// TIA Portal V20 export
Screen "Robot_PLP_Kuka"  1276x673
  ScreenItem "Zone01" at 710,47 size 522x643  Type=HmiGraphicView
  ScreenItem "Rectangle TG Control" at 241,104 size 465x354  Type=HmiRectangle
  ScreenItem "permanentareaborderrectangle" at 0,0 size 0x0  Type=HmiRectangle
  ScreenItem "Line_Header_X0_Y64" at 0,64 size 1280x0  Type=HmiLine
  ScreenItem "nbgMessages" at 19,459 size 687x203  Type=HmiAlarmControl
  ScreenItem "Button_Back" at 2,2 size 90x60  Type=HmiButton
  ScreenItem "Rectangle Robot Status" at 19,104 size 222x354  Type=HmiRectangle
  ScreenItem "Text Filed E- Stop" at 129,207 size 100x21  Type=HmiTextBox
  ScreenItem "Text Field In Auto On" at 24,138 size 100x21  Type=HmiTextBox
  ScreenItem "Text Field Home Position" at 24,161 size 100x21  Type=HmiTextBox
  ScreenItem "Text field PLP Status" at 19,103 size 222x31  Type=HmiTextBox
  ScreenItem "Text Field Manual" at 129,138 size 100x21  Type=HmiTextBox
  ScreenItem "Text Field System Ready" at 24,184 size 100x21  Type=HmiTextBox
  ScreenItem "Text Field Motor On" at 24,207 size 100x21  Type=HmiTextBox
  ScreenItem "Text Field In Cycle" at 24,230 size 100x21  Type=HmiTextBox
  ScreenItem "Text Field Cycle On" at 24,253 size 100x21  Type=HmiTextBox
  ScreenItem "Text Field On Path" at 24,276 size 100x21  Type=HmiTextBox
  ScreenItem "Text Field ProgNumReq" at 24,299 size 100x21  Type=HmiTextBox
  ScreenItem "Text Field Task OK" at 24,322 size 100x21  Type=HmiTextBox
  ScreenItem "Text Field Tryout Mode" at 129,161 size 100x21  Type=HmiTextBox
  ScreenItem "Text Field Stop" at 129,184 size 100x21  Type=HmiTextBox
  ScreenItem "Text Filed Error" at 129,230 size 100x21  Type=HmiTextBox
  ScreenItem "IO Field Feedback Program" at 129,280 size 100x21  Type=HmiIOField
  ScreenItem "Text Field Feedback Program" at 134,250 size 89x30  Type=HmiTextBox
  ScreenItem "Text Field In Home Pos" at 24,345 size 100x21  Type=HmiTextBox
  ScreenItem "Text Field In Work Pos" at 24,368 size 100x21  Type=HmiTextBox
  ScreenItem "Text Field In Pounce Pos" at 24,391 size 100x21  Type=HmiTextBox
  ScreenItem "Rectangle Clear Style" at 251,262 size 85x56  Type=HmiRectangle
  ScreenItem "Button Clear Style" at 252,263 size 83x54  Type=HmiButton
  ScreenItem "Clear Style Interlock" at 0,0 size 100x30  Type=HmiCircle
  ScreenItem "Rectangle Select Style1" at 251,140 size 85x56  Type=HmiRectangle
  ScreenItem "Button Select Style1" at 252,141 size 83x54  Type=HmiButton
  ScreenItem "Select Style Interlock1" at 0,0 size 100x30  Type=HmiCircle
  ScreenItem "Rectangle Select Style2" at 341,140 size 85x56  Type=HmiRectangle
  ScreenItem "Button Select Style2" at 342,141 size 83x54  Type=HmiButton
  ScreenItem "Select Style Interlock2" at 0,0 size 100x30  Type=HmiCircle
  ScreenItem "Rectangle Select Style3" at 431,140 size 85x56  Type=HmiRectangle
  ScreenItem "Button Select Style3" at 432,141 size 83x54  Type=HmiButton
  ScreenItem "Select Style Interlock3" at 0,0 size 100x30  Type=HmiCircle
  ScreenItem "Rectangle Select Style4" at 521,140 size 85x56  Type=HmiRectangle
  ScreenItem "Button Select Style4" at 522,141 size 83x54  Type=HmiButton
  ScreenItem "Select Style Interlock4" at 0,0 size 100x30  Type=HmiCircle
  ScreenItem "Rectangle Select Style5" at 611,140 size 85x56  Type=HmiRectangle
  ScreenItem "Button Select Style5" at 612,141 size 83x54  Type=HmiButton
  ScreenItem "Select Style Interlock5" at 0,0 size 100x30  Type=HmiCircle
  ScreenItem "Rectangle Select Style6" at 251,201 size 85x56  Type=HmiRectangle
  ScreenItem "Button Select Style6" at 252,202 size 83x54  Type=HmiButton
  ScreenItem "Select Style Interlock6" at 0,0 size 100x30  Type=HmiCircle
  ScreenItem "Rectangle Select Style7" at 341,201 size 85x56  Type=HmiRectangle
  ScreenItem "Button Select Style7" at 342,202 size 83x54  Type=HmiButton
  ScreenItem "Select Style Interlock7" at 0,0 size 100x30  Type=HmiCircle
  ScreenItem "Rectangle Select Style8" at 431,201 size 85x56  Type=HmiRectangle
  ScreenItem "Button Select Style8" at 432,202 size 83x54  Type=HmiButton
  ScreenItem "Select Style Interlock8" at 0,0 size 100x30  Type=HmiCircle
  ScreenItem "Rectangle Select Style9" at 521,201 size 85x56  Type=HmiRectangle
  ScreenItem "Button Select Style9" at 522,202 size 83x54  Type=HmiButton
  ScreenItem "Select Style Interlock9" at 0,0 size 100x30  Type=HmiCircle
  ScreenItem "Rectangle Select Style10" at 611,201 size 85x56  Type=HmiRectangle
  ScreenItem "Button Select Style10" at 612,202 size 83x54  Type=HmiButton
  ScreenItem "Select Style Interlock10" at 0,0 size 100x30  Type=HmiCircle
  ScreenItem "Rectangle Go Home" at 251,380 size 85x56  Type=HmiRectangle
  ScreenItem "Button Go Home" at 252,381 size 83x54  Type=HmiButton
  ScreenItem "Go Home Interlock" at 0,0 size 100x30  Type=HmiCircle
  ScreenItem "Rectangle Go Work" at 341,380 size 85x56  Type=HmiRectangle
  ScreenItem "Button Go Work" at 342,381 size 83x54  Type=HmiButton
  ScreenItem "Go Work Interlock" at 0,0 size 100x30  Type=HmiCircle
  ScreenItem "Rectangle Go Pounce" at 431,380 size 85x56  Type=HmiRectangle
  ScreenItem "Button Go Pounce" at 432,381 size 83x54  Type=HmiButton
  ScreenItem "Go Pounce Interlock" at 0,0 size 100x30  Type=HmiCircle
  ScreenItem "Text field Select Style" at 241,103 size 465x31  Type=HmiTextBox
  ScreenItem "Text field TG Control" at 241,335 size 465x31  Type=HmiTextBox
  ScreenItem "Text Field To Home Pos" at 129,345 size 100x21  Type=HmiTextBox
  ScreenItem "Text Field To Work Pos" at 129,368 size 100x21  Type=HmiTextBox
  ScreenItem "Text Field To Pounce Pos" at 129,391 size 100x21  Type=HmiTextBox
  ScreenItem "Rectangle TG1_4" at 40,0 size 185x55  Type=HmiRectangle
  ScreenItem "Rectangle TGC_4" at 0,0 size 40x55  Type=HmiRectangle
  ScreenItem "Text field TG1 Status_4" at 2,17 size 36x21  Type=HmiTextBox
  ScreenItem "Text Field TG5 In Pounce Pos" at 43,28 size 90x21  Type=HmiTextBox
  ScreenItem "Text Field TG5 In Work Pos" at 132,28 size 90x21  Type=HmiTextBox
  ScreenItem "Text Field TG5 Fault" at 43,6 size 90x21  Type=HmiTextBox
  ScreenItem "Text Field TG5 In Home Pos" at 132,6 size 90x21  Type=HmiTextBox
  ScreenItem "Rectangle TG1_5" at 40,0 size 185x55  Type=HmiRectangle
  ScreenItem "Rectangle TGC_5" at 0,0 size 40x55  Type=HmiRectangle
  ScreenItem "Text field TG1 Status_5" at 2,17 size 36x21  Type=HmiTextBox
  ScreenItem "Text Field TG6 In Pounce Pos" at 43,28 size 90x21  Type=HmiTextBox
  ScreenItem "Text Field TG6 In Work Pos" at 132,28 size 90x21  Type=HmiTextBox
  ScreenItem "Text Field TG6 Fault" at 43,6 size 90x21  Type=HmiTextBox
  ScreenItem "Text Field TG6 In Home Pos" at 132,6 size 90x21  Type=HmiTextBox
  ScreenItem "Rectangle TG1_6" at 40,0 size 185x55  Type=HmiRectangle
  ScreenItem "Rectangle TGC_6" at 0,0 size 40x55  Type=HmiRectangle
  ScreenItem "Text field TG1 Status_6" at 2,17 size 36x21  Type=HmiTextBox
  ScreenItem "Text Field TG7 In Pounce Pos" at 43,28 size 90x21  Type=HmiTextBox
  ScreenItem "Text Field TG7 In Work Pos" at 132,28 size 90x21  Type=HmiTextBox
  ScreenItem "Text Field TG7 Fault" at 43,6 size 90x21  Type=HmiTextBox
  ScreenItem "Text Field TG7 In Home Pos" at 132,6 size 90x21  Type=HmiTextBox
  ScreenItem "Rectangle TG1_7" at 40,0 size 185x55  Type=HmiRectangle
  ScreenItem "Rectangle TGC_7" at 0,0 size 40x55  Type=HmiRectangle
  ScreenItem "Text field TG1 Status_7" at 2,17 size 36x21  Type=HmiTextBox
  ScreenItem "Text Field TG8 In Pounce Pos" at 43,28 size 90x21  Type=HmiTextBox
  ScreenItem "Text Field TG8 In Work Pos" at 132,28 size 90x21  Type=HmiTextBox
  ScreenItem "Text Field TG8 Fault" at 43,6 size 90x21  Type=HmiTextBox
  ScreenItem "Text Field TG8 In Home Pos" at 132,6 size 90x21  Type=HmiTextBox
  ScreenItem "Rectangle TG1" at 40,0 size 185x55  Type=HmiRectangle
  ScreenItem "Rectangle TGC" at 0,0 size 40x55  Type=HmiRectangle
  ScreenItem "Text field TG1 Status" at 2,17 size 36x21  Type=HmiTextBox
  ScreenItem "Text Field TG1 In Pounce Pos" at 43,28 size 90x21  Type=HmiTextBox
  ScreenItem "Text Field TG1 In Work Pos" at 132,28 size 90x21  Type=HmiTextBox
  ScreenItem "Text Field TG1 Fault" at 43,6 size 90x21  Type=HmiTextBox
  ScreenItem "Text Field TG1 In Home Pos" at 132,6 size 90x21  Type=HmiTextBox
  ScreenItem "Select NC Locator" at 403,64 size 290x37  Type=HmiSymbolicIOField
  ScreenItem "Title_ScreenOverview_X390_Y2_3" at 384,5 size 510x57  Type=HmiTextBox
